Fanuc KAREL source: kd00043.KL

-- PROVISIONAL review KL for V1013-1; original PC SHA256 068e518ae42fb82ff33390cdc1c10c01b1df6d4a3f948b92936ae0e02fbb5567
-- Incomplete behavior may be omitted. Consult companion uncertainty JSON. Do not deploy.
PROGRAM KD00043
%NOLOCKGROUP
VAR
  I : INTEGER
  J : INTEGER
  B : BOOLEAN
  R : REAL
  S : STRING[80]
-- UNRESOLVED_DECL C type=000014
BEGIN
  -- UNRESOLVED_PC offsets 5-12; opcodes 9D,23
  -- UNRESOLVED_PC offsets 17-21; opcodes 7F
END KD00043
